(* IEC 61131-3 sources: nautilus/website/lessons/b1-blink/solution, 1 file *)

(* ---- program.st ---- *)
PROGRAM Blink
VAR
    tick : TON;   (* counts half a second, then says so for one scan *)
END_VAR

tick(IN := NOT tick.Q, PT := T#500ms);

IF tick.Q THEN
    Lamp := NOT Lamp;
END_IF;
END_PROGRAM
